Fanuc KAREL source: kt00244.KL

-- PROVISIONAL review KL for V940-1; original PC SHA256 8c773435d6b352c168c2e6db0eefce32e450a2faa25729cefd7fbdb17c67a096
-- Incomplete behavior may be omitted. Consult companion uncertainty JSON. Do not deploy.
PROGRAM KT00244
%NOLOCKGROUP
VAR
  I2 : INTEGER
  OUT : INTEGER
-- UNRESOLVED_DECL Y1 type=002018
BEGIN
  -- V9_ZERO_TABLE_METADATA_HINT layout=0001; no indexed target words; source/name/runtime held
  -- UNRESOLVED_PC offsets 5-19; opcodes 2E,22,9D,33,B2
  -- UNRESOLVED_PC offsets 24-35; opcodes 2E,23
  -- UNRESOLVED_PC offsets 40-62; opcodes 22,9D,33,B1,21,47,23
  -- UNRESOLVED_PC offsets 67-71; opcodes 7F
END KT00244
